Staubli VAL3: utCommon.dtx

public bool bDisabled
public string sText
public string sID
public string sPage
